(* IEC 61131-3 sources: codesys-ai-industrial-robot-control/plc/src/Process, 4 files *)

(* ---- F_SelectBin.st ---- *)
(*
    F_SelectBin
    Purpose : Bin selection of spec section 7.2:
              1. no valid vision, low confidence, or an AI decision saying the identification
                 is unreliable -> Quarantine
              2. quality Scrap -> Scrap, quality Rework -> Rework
              3. otherwise the type bin of the detected class
*)
FUNCTION F_SelectBin : E_Bin
VAR_INPUT
    stRec : ST_PartRecord;
    rConfThreshold : REAL;
    aClassToBin : ARRAY[0..2] OF E_Bin;
END_VAR

IF NOT stRec.xVisionValid OR stRec.rConfidence < rConfThreshold THEN
    F_SelectBin := E_Bin.Quarantine;
ELSIF stRec.eDecisionSource = E_DecisionSource.Ai AND NOT stRec.xIdentReliable THEN
    F_SelectBin := E_Bin.Quarantine;
ELSIF stRec.eQuality = E_Quality.Scrap THEN
    F_SelectBin := E_Bin.Scrap;
ELSIF stRec.eQuality = E_Quality.Rework THEN
    F_SelectBin := E_Bin.Rework;
ELSIF stRec.usiClass <= 2 THEN
    F_SelectBin := aClassToBin[stRec.usiClass];
ELSE
    F_SelectBin := E_Bin.Quarantine;
END_IF

(* ---- FB_PartTracker.st ---- *)
(*
    FB_PartTracker
    Purpose : Tracks every part from the PE1 capture until it is placed, missed or dropped.
              Applies vision and decision messages (only for known part ids, each message once),
              falls back to the rule-based decision at GVL_Params.tDecisionDeadline and marks
              parts that leave the pick window as missed.
    Inputs  : lrBeltPos [mm], xPE1Rising, stVision, stDecision, itfAlarms, xDecisionActive
    Outputs : stCapture (capture request to the vision service), udiPlaced/udiMissed/udiDropped,
              udiVisionMsgs (vision results applied)
    Methods : NextPickable, FindPart, GetRecord, SetState, CurrentX; property Count
    Belt X  : current X of a part = lrX (belt frame at capture) + (lrBeltPos - lrBeltPosAtCapture)
    Alarms  : QueueOverflow (condition: raised while full, cleared on the next successful capture);
              DecisionFallback, VisionMissing, LowConfidence, PartMissed (one-shot events)
*)
FUNCTION_BLOCK FB_PartTracker
VAR_INPUT
    lrBeltPos : LREAL;
    xPE1Rising : BOOL;
    stVision : ST_VisionMsg;
    stDecision : ST_DecisionMsg;
    itfAlarms : I_AlarmSink;
    // TRUE: an AI decision service answers (bridge); FALSE: the rule decides a part as soon as
    // vision has identified it, without waiting for the deadline and without DecisionFallback
    xDecisionActive : BOOL := TRUE;
END_VAR
VAR_OUTPUT
    stCapture : ST_CaptureMsg;
    udiPlaced : UDINT;
    udiMissed : UDINT;
    udiDropped : UDINT;
    udiVisionMsgs : UDINT;
END_VAR
VAR
    fbQueue : FB_PartQueue;
    fbTrigger : FB_CameraTrigger;
    fbIntake : FB_MessageIntake;
    stRec : ST_PartRecord;
    stNew : ST_PartRecord;
    uiIdx : UINT;
    i : UINT;
END_VAR

// 1. New part at the camera photo-eye.
fbTrigger(xPE1Rising := xPE1Rising, lrBeltPos := lrBeltPos);
stCapture := fbTrigger.stCapture;
IF fbTrigger.xNewPart THEN
    stRec := stNew;
    stRec.udiPartId := fbTrigger.udiNewPartId;
    stRec.lrBeltPosAtCapture := lrBeltPos;
    stRec.lrX := GVL_CellGeometry.PE1_X;         // until vision reports the exact position
    stRec.eState := E_PartState.Captured;
    stRec.tCaptured := TIME();
    IF fbQueue.AddRecord(stRec) = 0 THEN
        RaiseAlarm(E_AlarmId.QueueOverflow);
    ELSIF itfAlarms <> 0 THEN
        itfAlarms.Clear(E_AlarmId.QueueOverflow);
    END_IF
END_IF

// 2. Messages from the bridge (each sequence number once, known part ids only).
fbIntake(stVision := stVision, stDecision := stDecision);
IF fbIntake.xVisionNew THEN
    uiIdx := fbQueue.FindIndex(stVision.udiPartId);
    IF uiIdx > 0 THEN
        stRec := fbQueue.GetRecord(uiIdx);
        IF stRec.eState = E_PartState.Captured THEN
            stRec.xVisionValid := stVision.xValid;
            stRec.usiClass := stVision.usiClass;
            stRec.rConfidence := stVision.rConfidence;
            stRec.lrX := stVision.lrX;
            stRec.lrY := stVision.lrY;
            stRec.lrTheta := stVision.lrTheta;
            stRec.eState := E_PartState.Identified;
            fbQueue.PutRecord(uiIdx, stRec);
            udiVisionMsgs := udiVisionMsgs + 1;
            IF NOT xDecisionActive AND stRec.xVisionValid THEN
                stRec.eDecisionSource := E_DecisionSource.Fallback;
                stRec.eQuality := E_Quality.Unknown;
                Decide(uiIdx, stRec);
            END_IF
        END_IF
    END_IF
END_IF
IF fbIntake.xDecisionNew THEN
    uiIdx := fbQueue.FindIndex(stDecision.udiPartId);
    IF uiIdx > 0 THEN
        stRec := fbQueue.GetRecord(uiIdx);
        IF stRec.eState = E_PartState.Identified THEN
            stRec.eQuality := stDecision.eQuality;
            stRec.rQualityProb := stDecision.rQualityProb;
            stRec.xIdentReliable := stDecision.xIdentReliable;
            stRec.eDecisionSource := E_DecisionSource.Ai;
            Decide(uiIdx, stRec);
        END_IF
    END_IF
END_IF

// 3. Deadline fallback and parts leaving the pick window.
FOR i := 1 TO GVL_Config.MAX_PARTS DO
    stRec := fbQueue.GetRecord(i);
    IF (stRec.eState = E_PartState.Captured OR stRec.eState = E_PartState.Identified)
       AND TIME() - stRec.tCaptured >= GVL_Params.tDecisionDeadline THEN
        stRec.eDecisionSource := E_DecisionSource.Fallback;
        stRec.eQuality := E_Quality.Unknown;
        IF NOT stRec.xVisionValid THEN
            RaiseEventAlarm(E_AlarmId.VisionMissing);
        END_IF
        IF xDecisionActive THEN
            RaiseEventAlarm(E_AlarmId.DecisionFallback);
        END_IF
        Decide(i, stRec);
        stRec := fbQueue.GetRecord(i);
    END_IF
    IF (stRec.eState = E_PartState.Captured OR stRec.eState = E_PartState.Identified
        OR stRec.eState = E_PartState.Decided)
       AND CurrentX(i) > GVL_CellGeometry.PICK_WINDOW_END_X THEN
        SetState(i, E_PartState.Missed);
    END_IF
END_FOR

(* ---- FB_PickSequence.st ---- *)
(*
    FB_PickSequence
    Purpose : Pick-and-place cycle from the moving conveyor:
              home -> ready pose -> wait for a decided part in the pick window ->
              MC_TrackConveyorBelt (PCS_1 follows the part) -> linear approach / descend ->
              vacuum grip -> linear lift -> PTP to the target bin -> release -> retract.
    In/Out  : AxisGroup, ConveyorAxis, Robot (FB_Robot), Gripper (FB_VacuumGripper),
              Tracker (FB_PartTracker). The owner calls Robot, Gripper and Tracker each cycle.
    Inputs  : xRun - work on parts (FALSE: finish the current part, then go home and idle)
              xAbort - controlled stop now; the vacuum stays as it is (no dropped part)
              xReset - leave Error / Aborted to Idle. A part still held is placed in the
                       Quarantine bin on the next run; a scheduled part is marked missed.
    Outputs : eStep, xIdleAtHome, xBusy, udiPicked, udiPlaced, eLastBin, xPlacedPulse (one cycle)
    Errors  : every error first stops the robot (Aborting), then rests in Error.
    Window  : a pick is abandoned (part missed) if the part passes the pick window end before
              it is gripped.
    Moves   : linear only for the short tracked moves (PCS_1); PTP for long transfers, which
              avoids wrist/base singularities on Cartesian paths across the cell.
    Heights : approach, grip and lift heights follow the scheduled part's class
              (GVL_CellGeometry.PART_HEIGHTS).
*)
FUNCTION_BLOCK FB_PickSequence
VAR_IN_OUT
    AxisGroup : AXIS_GROUP_REF_SM3;
    ConveyorAxis : AXIS_REF_SM3;
    Robot : FB_Robot;
    Gripper : FB_VacuumGripper;
    Tracker : FB_PartTracker;
END_VAR
VAR_INPUT
    xRun : BOOL;
    xAbort : BOOL;
    xReset : BOOL;
END_VAR
VAR_OUTPUT
    eStep : E_PickStep;
    xIdleAtHome : BOOL;
    xBusy : BOOL;
    udiPicked : UDINT;
    udiPlaced : UDINT;
    eLastBin : E_Bin;
    xPlacedPulse : BOOL;
END_VAR
VAR
    fbTrack : MC_TrackConveyorBelt;
    tonRelease : TON;
    xTrackExec : BOOL;
    uiIdx : UINT;                       // slot of the part being handled, 0 = none
    stPart : ST_PartRecord;
    stObject : MC_COORD_REF;
    stTarget : SMC_POS_REF;
    stHeld : ST_PartRecord;
    xAtHome : BOOL;
    xFaultPending : BOOL;               // Aborting was entered because of an error
    xRecover : BOOL;                    // a held part must go to quarantine on the next run
    // robot command handshake
    iCmdPhase : INT;
    xRequested : BOOL;
    eReqCmd : E_RobotCmd;
    stReqTarget : SMC_POS_REF;
    xCmdDone : BOOL;
    xCmdError : BOOL;
    lrPartHeight : LREAL;               // grip height of the scheduled part's class [mm]
END_VAR
VAR CONSTANT
    RELEASE_TIME : TIME := T#200MS;      // vacuum off before retracting
END_VAR

xPlacedPulse := FALSE;
xCmdDone := FALSE;
xCmdError := FALSE;

// Robot command handshake: new command -> Execute FALSE -> TRUE -> wait for Done / Error.
CASE iCmdPhase OF
    1:
        Robot.eCmd := eReqCmd;
        Robot.stTarget := stReqTarget;
        Robot.xExecute := FALSE;
        iCmdPhase := 2;
    2:
        Robot.xExecute := TRUE;
        iCmdPhase := 3;
    3:
        IF Robot.xDone THEN
            Robot.xExecute := FALSE;
            iCmdPhase := 0;
            xCmdDone := TRUE;
        ELSIF Robot.xError THEN
            Robot.xExecute := FALSE;
            iCmdPhase := 0;
            xCmdError := TRUE;
        END_IF
END_CASE

fbTrack(AxisGroup := AxisGroup,
        ConveyorBelt := ConveyorAxis,
        Execute := xTrackExec,
        ConveyorBeltOrigin := GVL_CellGeometry.BELT_ORIGIN,
        InitialObjectPosition := stObject,
        CoordSystem := SMC_COORD_SYSTEM.PCS_1);

IF xAbort AND eStep <> E_PickStep.Idle AND eStep <> E_PickStep.Aborting
   AND eStep <> E_PickStep.Aborted AND eStep <> E_PickStep.Error THEN
    eStep := E_PickStep.Aborting;
    iCmdPhase := 0;
    xRequested := FALSE;
END_IF
IF xReset AND (eStep = E_PickStep.Error OR eStep = E_PickStep.Aborted) THEN
    IF Gripper.xHolding AND uiIdx > 0 THEN
        stPart.eTargetBin := E_Bin.Quarantine;       // unknown history: quarantine it
        xRecover := TRUE;
    ELSE
        Gripper.xCmdVacuum := FALSE;
        xRecover := FALSE;
        IF uiIdx > 0 THEN
            stHeld := Tracker.GetRecord(uiIdx);
            IF stHeld.eState = E_PartState.Scheduled OR stHeld.eState = E_PartState.Picked THEN
                Tracker.SetState(uiIdx, E_PartState.Missed);
            END_IF
            uiIdx := 0;
        END_IF
    END_IF
    eStep := E_PickStep.Idle;
    iCmdPhase := 0;
    xRequested := FALSE;
    xTrackExec := FALSE;
    xAtHome := FALSE;
    xFaultPending := FALSE;
    Robot.xExecute := FALSE;
END_IF

CASE eStep OF
    E_PickStep.Idle:
        IF xRun THEN
            IF xRecover THEN
                NextStep(E_PickStep.RecoverLift);   // a part is on the cup: straight up first
            ELSE
                NextStep(E_PickStep.MoveHome);
            END_IF
        END_IF

    E_PickStep.MoveHome:
        Request(E_RobotCmd.MovePtpAcs, GVL_CellGeometry.HOME_ACS);
        IF xCmdDone THEN
            xAtHome := TRUE;
            IF xRun THEN
                NextStep(E_PickStep.MoveReady);
            ELSE
                NextStep(E_PickStep.Idle);
            END_IF
        END_IF

    E_PickStep.RecoverLift:
        // after an abort the arm may stand anywhere (near the belt, a bin wall): lift vertically
        // to the ready height before any point-to-point move, whose path is not known
        stTarget := Robot.stActMcs;
        stTarget.c.Z := MAX(Robot.stActMcs.c.Z, GVL_CellGeometry.READY_POSE.Z);
        Request(E_RobotCmd.MoveLinMcs, stTarget);
        IF xCmdDone THEN
            NextStep(E_PickStep.MoveReady);
        END_IF

    E_PickStep.MoveReady:
        stTarget.c := GVL_CellGeometry.READY_POSE;
        Request(E_RobotCmd.MovePtpMcs, stTarget);
        IF xCmdDone THEN
            xAtHome := FALSE;
            IF xRecover THEN
                NextStep(E_PickStep.MoveToBin);     // the held part goes to its bin from Ready
            ELSE
                NextStep(E_PickStep.WaitPart);
            END_IF
        END_IF

    E_PickStep.WaitPart:
        IF NOT xRun THEN
            NextStep(E_PickStep.MoveHome);
        ELSE
            uiIdx := Tracker.NextPickable(GVL_CellGeometry.PE2_X,
                                          GVL_CellGeometry.PICK_WINDOW_END_X - GVL_CellGeometry.PICK_MARGIN);
            IF uiIdx > 0 THEN
                stPart := Tracker.GetRecord(uiIdx);
                lrPartHeight := GVL_CellGeometry.PART_HEIGHTS[MIN(stPart.usiClass, 2)];
                stObject.X := Tracker.CurrentX(uiIdx);
                stObject.Y := stPart.lrY;
                stObject.Z := GVL_CellGeometry.BELT_SURFACE_Z;
                stObject.A := stPart.lrTheta;
                stObject.B := 0;
                stObject.C := 0;
                Tracker.SetState(uiIdx, E_PartState.Scheduled);
                xTrackExec := FALSE;
                NextStep(E_PickStep.StartTracking);
            END_IF
        END_IF

    E_PickStep.StartTracking:
        xTrackExec := TRUE;
        IF fbTrack.Done THEN
            NextStep(E_PickStep.Approach);
        ELSIF fbTrack.Error THEN
            GoError();
        END_IF

    E_PickStep.Approach:
        Request(E_RobotCmd.MoveLinPcs1, TrackedPose(lrPartHeight + GVL_Params.lrApproachHeight));
        IF xCmdDone THEN
            NextStep(E_PickStep.Descend);
        END_IF

    E_PickStep.Descend:
        Request(E_RobotCmd.MoveLinPcs1, TrackedPose(lrPartHeight - GVL_Params.lrPickDepth));
        IF xCmdDone THEN
            NextStep(E_PickStep.Grip);
        END_IF

    E_PickStep.Grip:
        Gripper.xCmdVacuum := TRUE;
        IF Gripper.xHolding THEN
            Tracker.SetState(uiIdx, E_PartState.Picked);
            udiPicked := udiPicked + 1;
            NextStep(E_PickStep.Lift);
        ELSIF Gripper.HasError THEN
            Gripper.xCmdVacuum := FALSE;          // nothing is held
            Tracker.SetState(uiIdx, E_PartState.Dropped);
            uiIdx := 0;
            GoError();
        END_IF

    E_PickStep.Lift:
        Request(E_RobotCmd.MoveLinPcs1, TrackedPose(lrPartHeight + GVL_Params.lrApproachHeight));
        IF xCmdDone THEN
            xTrackExec := FALSE;
            NextStep(E_PickStep.MoveToBin);
        END_IF

    E_PickStep.MoveToBin:
        stTarget.c := GVL_CellGeometry.BIN_DROP[stPart.eTargetBin];
        Request(E_RobotCmd.MovePtpMcs, stTarget);
        IF xCmdDone THEN
            NextStep(E_PickStep.Release);
        END_IF

    E_PickStep.Release:
        Gripper.xCmdVacuum := FALSE;
        tonRelease(IN := TRUE, PT := RELEASE_TIME);
        IF tonRelease.Q THEN
            Tracker.SetState(uiIdx, E_PartState.Placed);
            uiIdx := 0;
            xRecover := FALSE;
            udiPlaced := udiPlaced + 1;
            eLastBin := stPart.eTargetBin;
            xPlacedPulse := TRUE;
            NextStep(E_PickStep.Retract);
        END_IF

    E_PickStep.Retract:
        stTarget.c := GVL_CellGeometry.BIN_DROP[stPart.eTargetBin];
        stTarget.c.Z := stTarget.c.Z + GVL_CellGeometry.RETRACT_HEIGHT;
        Request(E_RobotCmd.MoveLinMcs, stTarget);
        IF xCmdDone THEN
            IF xRun THEN
                NextStep(E_PickStep.MoveReady);
            ELSE
                NextStep(E_PickStep.MoveHome);
            END_IF
        END_IF

    E_PickStep.Aborting:
        Request(E_RobotCmd.Stop, stTarget);
        IF xCmdDone OR xCmdError THEN
            xTrackExec := FALSE;
            IF xFaultPending THEN
                xFaultPending := FALSE;
                NextStep(E_PickStep.Error);
            ELSE
                NextStep(E_PickStep.Aborted);
            END_IF
        END_IF

    E_PickStep.Aborted, E_PickStep.Error:
        ;   // wait for xReset
END_CASE

// The part passed the pick window end before it was gripped: give it up, do not chase it.
IF (eStep = E_PickStep.StartTracking OR eStep = E_PickStep.Approach OR eStep = E_PickStep.Descend
    OR eStep = E_PickStep.Grip) AND uiIdx > 0 AND NOT Gripper.xHolding
   AND Tracker.CurrentX(uiIdx) > GVL_CellGeometry.PICK_WINDOW_END_X THEN
    Gripper.xCmdVacuum := FALSE;
    Tracker.SetState(uiIdx, E_PartState.Missed);
    uiIdx := 0;
    xTrackExec := FALSE;
    iCmdPhase := 0;
    Robot.xExecute := FALSE;
    NextStep(E_PickStep.MoveReady);
END_IF

// A part lost while carrying it: stop the robot; the valve stays on (spec 5.4: no release outside
// a bin), Stopping / recovery decide what happens next.
IF (eStep = E_PickStep.Lift OR eStep = E_PickStep.MoveToBin) AND Gripper.HasError THEN
    Tracker.SetState(uiIdx, E_PartState.Dropped);
    uiIdx := 0;
    GoError();
END_IF
IF xCmdError AND eStep <> E_PickStep.Aborting AND eStep <> E_PickStep.Aborted
   AND eStep <> E_PickStep.Error THEN
    GoError();
END_IF

xIdleAtHome := eStep = E_PickStep.Idle AND xAtHome;
xBusy := eStep <> E_PickStep.Idle AND eStep <> E_PickStep.WaitPart
         AND eStep <> E_PickStep.Aborted AND eStep <> E_PickStep.Error;

(* ---- FB_SortingCell.st ---- *)
(*
    FB_SortingCell
    Purpose : The sorting cell as one PackML unit. Owns all equipment and maps the PackML states
              to equipment actions; computes the interlocks.
    In/Out  : AxisGroup (AxisGroup_Robot), ConveyorAxis (Axis_Conveyor)
    Inputs  : operator commands (GVL_Hmi), sensors and messages (GVL_Bridge), xLoopback (feedback := setpoint)
    Outputs : setpoints, belt and vacuum to the bridge; eState, eMode, ePickStep, aActAcs;
              diagnostics (newest alarm, alarm classes, worst joint, following errors)
    States  : Resetting  - acknowledge alarms, reset equipment and the pick sequence, forget the
                           tracked parts; done when safe and fault-free
              Starting / Unholding / Unsuspending - robot home -> ready, conveyor at speed
                           (a part still on the cup is placed in quarantine first)
              Execute    - automatic: pick sequence runs; Manual: jogging
              Stopping / Holding / Suspending / Completing - finish the current part, go home;
                           done when the sequence rests, the robot and the belt stand still
              Aborting   - controlled stop, vacuum kept; Clearing - reset the sequence
    Interlocks: Critical alarm or not safe -> Abort; Error alarm -> Stop; any bin full -> Suspend,
              and Unsuspend automatically when that bin is emptied (not after an operator Suspend).
              Resetting and Clearing are not interrupted by the alarms they are clearing.
*)
FUNCTION_BLOCK FB_SortingCell
VAR_IN_OUT
    AxisGroup : AXIS_GROUP_REF_SM3;
    ConveyorAxis : AXIS_REF_SM3;
END_VAR
VAR_INPUT
    eCommand : E_PackMLCommand;
    eModeRequest : E_PackMLMode := E_PackMLMode.Production;
    xAlarmAck : BOOL;
    axJogPlus : ARRAY[1..6] OF BOOL;
    axJogMinus : ARRAY[1..6] OF BOOL;
    rOverride : REAL := 1.0;
    xHeartbeat : BOOL;
    aJointPosFb : ARRAY[1..6] OF LREAL;
    aJointTorqueFb : ARRAY[1..6] OF LREAL;
    udiFeedbackSeq : UDINT;
    udiFeedbackForSeq : UDINT;                // setpoint sample the joint feedback answers
    xPE1 : BOOL;
    xVacuumOk : BOOL;
    axBinFull : ARRAY[E_Bin.TypeA..E_Bin.Quarantine] OF BOOL;
    xDoorClosed : BOOL := TRUE;
    xEStopOk : BOOL := TRUE;
    stVision : ST_VisionMsg;
    stDecision : ST_DecisionMsg;
    xDecisionActive : BOOL;                  // an AI decision service answers (bridge)
    xLoopback : BOOL;
END_VAR
VAR_OUTPUT
    aJointPosSp : ARRAY[1..6] OF LREAL;
    lrBeltPos : LREAL;
    lrBeltVel : LREAL;
    xVacuumOn : BOOL;
    stCapture : ST_CaptureMsg;
    eState : E_PackMLState := E_PackMLState.Stopped;
    eMode : E_PackMLMode := E_PackMLMode.Production;
    ePickStep : E_PickStep;
    aActAcs : ARRAY[1..6] OF LREAL;
    udiSetpointSeq : UDINT;                   // +1 per cycle with every setpoint sample
    // diagnostics (bridge, HMI)
    eNewestAlarm : E_AlarmId;
    xAlarmError : BOOL;
    xAlarmCritical : BOOL;
    iWorstJoint : INT;
    aFollowingError : ARRAY[1..6] OF LREAL;   // [deg]
END_VAR
VAR
    fbSm : FB_PackMLStateMachine;
    fbAlarms : FB_AlarmHandler;
    fbSafety : FB_SafetyMonitor;
    fbConv : FB_Conveyor;
    fbRobot : FB_Robot;
    fbMon : FB_JointMonitor;
    fbTracker : FB_PartTracker;
    fbSeq : FB_PickSequence;
    fbVac : FB_VacuumGripper;
    aBins : ARRAY[E_Bin.TypeA..E_Bin.Quarantine] OF FB_Bin;
    fbPe1 : FB_PhotoEye;
    fbWatchdog : FB_BridgeWatchdog;
    fbJog : SMC_GroupJog2;
    eBin : E_Bin;
    i : INT;
    xAnyBinFull : BOOL;
    xSuspendedByBin : BOOL;             // the current suspension was caused by a full bin
    xComplete : BOOL;
    xAutoMode : BOOL;
    xRunBelt : BOOL;
    xJog : BOOL;
    xMotionStill : BOOL;                // pick sequence resting, robot and belt standing still
    lrSpeedFactor : LREAL;
    aFeedback : ARRAY[1..6] OF LREAL;
END_VAR
VAR CONSTANT
    REDUCED_SPEED_FACTOR : LREAL := 0.25;   // Maintenance mode and Manual with the door open
    JOG_VELOCITY : LREAL := 30;             // [deg/s] joint jog
    JOG_ACCELERATION : LREAL := 300;        // [deg/s2]
    JOG_JERK : LREAL := 3000;               // [deg/s3]
    JOG_MAX_LINEAR : LREAL := 100;          // [mm] per jog edge
    JOG_MAX_ANGULAR : LREAL := 45;          // [deg] per jog edge
    BELT_STANDSTILL : LREAL := 0.5;         // [mm/s] belt counts as stopped below this
END_VAR

eState := fbSm.eState;
eMode := fbSm.eMode;
xAutoMode := eMode <> E_PackMLMode.Manual;

fbRobot.itfAlarms := fbAlarms;
fbConv.itfAlarms := fbAlarms;
fbVac.itfAlarms := fbAlarms;
fbTracker.itfAlarms := fbAlarms;
fbSafety.itfAlarms := fbAlarms;
fbMon.itfAlarms := fbAlarms;
fbWatchdog.itfAlarms := fbAlarms;

// --- safety and alarm acknowledgement --------------------------------------------------------
fbSafety(xEStopOk := xEStopOk, xDoorClosed := xDoorClosed, eMode := eMode,
         xResetCmd := eState = E_PackMLState.Resetting OR eState = E_PackMLState.Clearing);
IF xAlarmAck OR (fbSm.xStateChanged AND (eState = E_PackMLState.Resetting OR eState = E_PackMLState.Clearing)) THEN
    fbAlarms.AcknowledgeAll();
END_IF

// --- bins --------------------------------------------------------------------------------------
xAnyBinFull := FALSE;
FOR eBin := E_Bin.TypeA TO E_Bin.Quarantine DO
    aBins[eBin](eBin := eBin,
                xFullSensor := axBinFull[eBin],
                xPlaced := fbSeq.xPlacedPulse AND fbSeq.eLastBin = eBin);
    xAnyBinFull := xAnyBinFull OR aBins[eBin].xFull;
END_FOR
IF xAnyBinFull THEN
    fbAlarms.Raise(E_AlarmId.BinFull);
ELSE
    fbAlarms.Clear(E_AlarmId.BinFull);
END_IF

// --- PackML state actions ----------------------------------------------------------------------
xComplete := FALSE;
xRunBelt := FALSE;
xJog := FALSE;
fbSeq.xRun := FALSE;
fbSeq.xAbort := FALSE;
fbSeq.xReset := FALSE;
xMotionStill := (fbSeq.eStep = E_PickStep.Idle OR fbSeq.eStep = E_PickStep.Error
                 OR fbSeq.eStep = E_PickStep.Aborted)
                AND NOT fbRobot.xMoving AND ABS(fbConv.lrActVelocity) < BELT_STANDSTILL;
CASE eState OF
    E_PackMLState.Resetting:
        fbSeq.xReset := TRUE;
        fbTracker.Clear();                        // parts on the belt are unknown after a stop
        fbRobot.Reset();
        fbVac.Reset();
        fbConv.Reset();
        xSuspendedByBin := FALSE;
        xComplete := fbSafety.xSafeToMove AND fbRobot.xReady AND fbSeq.eStep = E_PickStep.Idle
                     AND NOT fbAlarms.xCriticalActive AND NOT fbAlarms.xErrorActive;

    E_PackMLState.Starting, E_PackMLState.Unholding, E_PackMLState.Unsuspending:
        IF xAutoMode THEN
            fbSeq.xRun := TRUE;
            xRunBelt := TRUE;
            xComplete := fbSeq.eStep = E_PickStep.WaitPart AND fbConv.xAtSpeed;
        ELSE
            xComplete := fbRobot.xReady;
        END_IF

    E_PackMLState.Execute:
        xSuspendedByBin := xAnyBinFull;          // a full bin in Execute raises the suspension
        IF xAutoMode THEN
            fbSeq.xRun := TRUE;
            xRunBelt := TRUE;
        ELSE
            xJog := TRUE;
        END_IF

    E_PackMLState.Stopping, E_PackMLState.Holding, E_PackMLState.Suspending, E_PackMLState.Completing:
        xComplete := xMotionStill;

    E_PackMLState.Aborting:
        fbSeq.xAbort := TRUE;
        xComplete := NOT fbRobot.xMoving AND (fbSeq.eStep = E_PickStep.Aborted
                     OR fbSeq.eStep = E_PickStep.Idle OR fbSeq.eStep = E_PickStep.Error);

    E_PackMLState.Clearing:
        fbSeq.xReset := TRUE;
        fbRobot.Reset();
        fbVac.Reset();
        fbConv.Reset();
        xComplete := fbSafety.xSafeToMove AND fbSeq.eStep = E_PickStep.Idle
                     AND NOT fbAlarms.xCriticalActive;
END_CASE

// --- equipment ---------------------------------------------------------------------------------
IF eMode = E_PackMLMode.Maintenance OR fbSafety.xReducedSpeed THEN
    lrSpeedFactor := REDUCED_SPEED_FACTOR;
ELSE
    lrSpeedFactor := 1.0;
END_IF

fbPe1(xRaw := xPE1);
fbTracker(lrBeltPos := fbConv.lrPosition, xPE1Rising := fbPe1.xRising,
          stVision := stVision, stDecision := stDecision, xDecisionActive := xDecisionActive);
fbSeq(AxisGroup := AxisGroup, ConveyorAxis := ConveyorAxis,
      Robot := fbRobot, Gripper := fbVac, Tracker := fbTracker);
fbVac(xVacuumOk := xVacuumOk, tGripTimeout := GVL_Params.tVacuumTimeout);

fbRobot.xEnable := eState <> E_PackMLState.Stopped;
fbRobot.lrOverride := REAL_TO_LREAL(rOverride) * lrSpeedFactor;
fbRobot(AxisGroup := AxisGroup);

fbJog.Enable := xJog AND fbRobot.xReady AND fbSafety.xSafeToMove;
FOR i := 1 TO 6 DO
    fbJog.Forward[i - 1] := axJogPlus[i];
    fbJog.Backward[i - 1] := axJogMinus[i];
END_FOR
fbJog(AxisGroup := AxisGroup,
      CoordSystem := SMC_COORD_SYSTEM.ACS,
      MaxLinearDistance := JOG_MAX_LINEAR,
      MaxAngularDistance := JOG_MAX_ANGULAR,
      Velocity := JOG_VELOCITY,
      Acceleration := JOG_ACCELERATION,
      Deceleration := JOG_ACCELERATION,
      Jerk := JOG_JERK,
      VelFactor := lrSpeedFactor,
      AccFactor := 1.0,
      JerkFactor := 1.0);

fbConv(Axis := ConveyorAxis,
       xEnable := eState <> E_PackMLState.Stopped,
       lrVelocity := GVL_Params.lrBeltSpeed,
       xRun := xRunBelt AND fbSafety.xSafeToMove);

FOR i := 1 TO 6 DO
    IF xLoopback THEN
        aFeedback[i] := fbRobot.aSetAcs[i];
    ELSE
        aFeedback[i] := aJointPosFb[i];
    END_IF
END_FOR
udiSetpointSeq := udiSetpointSeq + 1;
fbMon(aSetpoint := fbRobot.aSetAcs, aFeedback := aFeedback, aTorque := aJointTorqueFb,
      udiFeedbackSeq := udiFeedbackSeq, udiSetpointSeq := udiSetpointSeq,
      udiFeedbackForSeq := udiFeedbackForSeq, xLoopback := xLoopback, xActive := fbRobot.xReady);
fbWatchdog(xHeartbeat := xHeartbeat, xEnable := NOT xLoopback AND eState <> E_PackMLState.Stopped);

// --- PackML ------------------------------------------------------------------------------------
fbAlarms();
fbSm(eCommand := eCommand,
     eModeRequest := eModeRequest,
     xStateComplete := xComplete,
     xAbortRequest := NOT fbSafety.xSafeToMove
                      OR (fbAlarms.xCriticalActive AND eState <> E_PackMLState.Resetting
                          AND eState <> E_PackMLState.Clearing),
     xStopRequest := fbAlarms.xErrorActive AND eState <> E_PackMLState.Resetting,
     xSuspendRequest := xAnyBinFull,
     xUnsuspendRequest := xSuspendedByBin AND NOT xAnyBinFull);

// --- outputs to the bridge ---------------------------------------------------------------------
aJointPosSp := fbRobot.aSetAcs;
lrBeltPos := fbConv.lrPosition;
lrBeltVel := fbConv.lrActVelocity;
xVacuumOn := fbVac.xValveOn;
stCapture := fbTracker.stCapture;
eState := fbSm.eState;
eMode := fbSm.eMode;
ePickStep := fbSeq.eStep;
eNewestAlarm := fbAlarms.eNewest;
xAlarmError := fbAlarms.xErrorActive;
xAlarmCritical := fbAlarms.xCriticalActive;
iWorstJoint := fbMon.iWorstJoint;
aFollowingError := fbMon.aFollowingError;
FOR i := 1 TO 6 DO
    CASE i OF
        1: aActAcs[i] := fbRobot.stActAcs.a.a0;
        2: aActAcs[i] := fbRobot.stActAcs.a.a1;
        3: aActAcs[i] := fbRobot.stActAcs.a.a2;
        4: aActAcs[i] := fbRobot.stActAcs.a.a3;
        5: aActAcs[i] := fbRobot.stActAcs.a.a4;
        6: aActAcs[i] := fbRobot.stActAcs.a.a5;
    END_CASE
END_FOR
